  movel([0.125319, -1.305667, -2.614786, -0.791936, 1.570796, 1.696115],accel_mss,speed_ms,0,blend_radius_m)
  movel([0.123866, -1.307460, -2.613698, -0.791230, 1.570796, 1.694663],accel_mss,speed_ms,0,blend_radius_m)
  movel([0.121238, -1.311144, -2.611452, -0.789794, 1.570796, 1.692034],accel_mss,speed_ms,0,blend_radius_m)
  movel([0.120065, -1.313039, -2.610289, -0.789062, 1.570796, 1.690862],accel_mss,speed_ms,0,blend_radius_m)
  movel([0.118018, -1.316931, -2.607885, -0.787572, 1.570796, 1.688814],accel_mss,speed_ms,0,blend_radius_m)
  movel([0.117145, -1.318934, -2.606641, -0.786814, 1.570796, 1.687942],accel_mss,speed_ms,0,blend_radius_m)
  movel([0.116379, -1.320970, -2.605370, -0.786048, 1.570796, 1.687175],accel_mss,speed_ms,0,blend_radius_m)
  movel([0.115454, -1.323887, -2.603541, -0.784961, 1.570796, 1.686251],accel_mss,speed_ms,0,blend_radius_m)
  movel([0.114703, -1.326797, -2.601704, -0.783888, 1.570796, 1.685499],accel_mss,speed_ms,0,blend_radius_m)
  movel([0.114117, -1.329682, -2.599872, -0.782835, 1.570796, 1.684914],accel_mss,speed_ms,0,blend_radius_m)
  movel([0.113685, -1.332534, -2.598050, -0.781805, 1.570796, 1.684482],accel_mss,speed_ms,0,blend_radius_m)
  movel([0.113406, -1.335329, -2.596253, -0.780807, 1.570796, 1.684202],accel_mss,speed_ms,0,blend_radius_m)
  movel([0.113271, -1.338054, -2.594492, -0.779843, 1.570796, 1.684068],accel_mss,speed_ms,0,blend_radius_m)
  movel([0.113272, -1.340695, -2.592775, -0.778919, 1.570796, 1.684069],accel_mss,speed_ms,0,blend_radius_m)
  movel([0.113405, -1.343237, -2.591113, -0.778039, 1.570796, 1.684201],accel_mss,speed_ms,0,blend_radius_m)
  movel([0.114874, -1.352772, -2.584802, -0.774815, 1.570796, 1.685670],accel_mss,speed_ms,0,blend_radius_m)
  movel([0.115989, -1.360388, -2.579670, -0.772330, 1.570796, 1.686785],accel_mss,speed_ms,0,blend_radius_m)
  movel([0.116017, -1.361138, -2.579161, -0.772090, 1.570796, 1.686813],accel_mss,speed_ms,0,blend_radius_m)
  movel([0.120926, -1.357802, -2.581422, -0.773165, 1.570796, 1.691723],accel_mss,speed_ms,0,blend_radius_m)
  movel([0.125997, -1.354721, -2.583496, -0.774171, 1.570796, 1.696793],accel_mss,speed_ms,0,blend_radius_m)
  movel([0.131197, -1.351900, -2.585385, -0.775105, 1.570796, 1.701994],accel_mss,speed_ms,0,blend_radius_m)
  movel([0.136489, -1.349339, -2.587089, -0.775961, 1.570796, 1.707286],accel_mss,speed_ms,0,blend_radius_m)
  movel([0.141835, -1.347047, -2.588606, -0.776735, 1.570796, 1.712632],accel_mss,speed_ms,0,blend_radius_m)
  movel([0.147200, -1.345021, -2.589942, -0.777426, 1.570796, 1.717996],accel_mss,speed_ms,0,blend_radius_m)
  movel([0.152545, -1.343268, -2.591093, -0.778028, 1.570796, 1.723342],accel_mss,speed_ms,0,blend_radius_m)
  movel([0.157833, -1.341785, -2.592064, -0.778541, 1.570796, 1.728629],accel_mss,speed_ms,0,blend_radius_m)
  movel([0.160299, -1.341216, -2.592435, -0.778738, 1.570796, 1.731096],accel_mss,speed_ms,0,blend_radius_m)
  movel([0.162784, -1.340774, -2.592724, -0.778892, 1.570796, 1.733580],accel_mss,speed_ms,0,blend_radius_m)
  movel([0.165263, -1.340467, -2.592923, -0.778998, 1.570796, 1.736060],accel_mss,speed_ms,0,blend_radius_m)
  movel([0.167711, -1.340305, -2.593029, -0.779055, 1.570796, 1.738507],accel_mss,speed_ms,0,blend_radius_m)
  movel([0.170105, -1.340295, -2.593036, -0.779058, 1.570796, 1.740901],accel_mss,speed_ms,0,blend_radius_m)
  movel([0.172421, -1.340447, -2.592937, -0.779005, 1.570796, 1.743217],accel_mss,speed_ms,0,blend_radius_m)
  movel([0.174636, -1.340766, -2.592729, -0.778894, 1.570796, 1.745433],accel_mss,speed_ms,0,blend_radius_m)
  movel([0.176726, -1.341259, -2.592407, -0.778723, 1.570796, 1.747522],accel_mss,speed_ms,0,blend_radius_m)
  movel([0.178667, -1.341936, -2.591965, -0.778488, 1.570796, 1.749464],accel_mss,speed_ms,0,blend_radius_m)
  movel([0.180439, -1.342801, -2.591399, -0.778189, 1.570796, 1.751235],accel_mss,speed_ms,0,blend_radius_m)
  movel([0.182015, -1.343863, -2.590703, -0.777823, 1.570796, 1.752811],accel_mss,speed_ms,0,blend_radius_m)
  movel([0.183374, -1.345125, -2.589873, -0.777390, 1.570796, 1.754170],accel_mss,speed_ms,0,blend_radius_m)
  movel([0.184492, -1.346595, -2.588905, -0.776889, 1.570796, 1.755289],accel_mss,speed_ms,0,blend_radius_m)
  movel([0.185353, -1.348277, -2.587793, -0.776319, 1.570796, 1.756149],accel_mss,speed_ms,0,blend_radius_m)
  movel([0.185931, -1.350176, -2.586533, -0.775680, 1.570796, 1.756728],accel_mss,speed_ms,0,blend_radius_m)
  movel([0.186205, -1.352297, -2.585119, -0.774972, 1.570796, 1.757002],accel_mss,speed_ms,0,blend_radius_m)
  movel([0.186151, -1.355276, -2.583124, -0.773989, 1.570796, 1.756947],accel_mss,speed_ms,0,blend_radius_m)
  movel([0.185726, -1.358424, -2.581001, -0.772963, 1.570796, 1.756523],accel_mss,speed_ms,0,blend_radius_m)
  movel([0.184990, -1.361689, -2.578786, -0.771914, 1.570796, 1.755786],accel_mss,speed_ms,0,blend_radius_m)
  movel([0.184002, -1.365022, -2.576509, -0.770858, 1.570796, 1.754798],accel_mss,speed_ms,0,blend_radius_m)
  movel([0.182819, -1.368372, -2.574204, -0.769813, 1.570796, 1.753615],accel_mss,speed_ms,0,blend_radius_m)
  movel([0.181495, -1.371694, -2.571903, -0.768792, 1.570796, 1.752291],accel_mss,speed_ms,0,blend_radius_m)
  movel([0.178658, -1.378063, -2.567448, -0.766878, 1.570796, 1.749455],accel_mss,speed_ms,0,blend_radius_m)
  movel([0.176687, -1.382024, -2.564648, -0.765716, 1.570796, 1.747483],accel_mss,speed_ms,0,blend_radius_m)
  movel([0.174549, -1.385880, -2.561901, -0.764608, 1.570796, 1.745346],accel_mss,speed_ms,0,blend_radius_m)
  movel([0.172265, -1.389646, -2.559198, -0.763545, 1.570796, 1.743062],accel_mss,speed_ms,0,blend_radius_m)
  movel([0.169850, -1.393345, -2.556522, -0.762522, 1.570796, 1.740646],accel_mss,speed_ms,0,blend_radius_m)
  movel([0.167323, -1.396990, -2.553866, -0.761533, 1.570796, 1.738120],accel_mss,speed_ms,0,blend_radius_m)
  movel([0.164703, -1.400600, -2.551217, -0.760572, 1.570796, 1.735499],accel_mss,speed_ms,0,blend_radius_m)
  movel([0.159243, -1.407786, -2.545886, -0.758717, 1.570796, 1.730039],accel_mss,speed_ms,0,blend_radius_m)
  movel([0.162416, -1.409703, -2.544451, -0.758235, 1.570796, 1.733213],accel_mss,speed_ms,0,blend_radius_m)
  movel([0.164019, -1.410829, -2.543606, -0.757954, 1.570796, 1.734815],accel_mss,speed_ms,0,blend_radius_m)
  movel([0.165312, -1.412098, -2.542651, -0.757640, 1.570796, 1.736108],accel_mss,speed_ms,0,blend_radius_m)
  movel([0.165766, -1.412796, -2.542125, -0.757468, 1.570796, 1.736562],accel_mss,speed_ms,0,blend_radius_m)
  movel([0.166050, -1.413541, -2.541562, -0.757286, 1.570796, 1.736847],accel_mss,speed_ms,0,blend_radius_m)
  movel([0.166139, -1.414334, -2.540963, -0.757092, 1.570796, 1.736935],accel_mss,speed_ms,0,blend_radius_m)
  movel([0.166002, -1.415178, -2.540323, -0.756887, 1.570796, 1.736798],accel_mss,speed_ms,0,blend_radius_m)
  movel([0.165610, -1.416074, -2.539643, -0.756671, 1.570796, 1.736406],accel_mss,speed_ms,0,blend_radius_m)
  movel([0.164930, -1.417031, -2.538917, -0.756442, 1.570796, 1.735726],accel_mss,speed_ms,0,blend_radius_m)
  movel([0.163937, -1.418049, -2.538141, -0.756199, 1.570796, 1.734733],accel_mss,speed_ms,0,blend_radius_m)
  movel([0.162601, -1.419130, -2.537317, -0.755943, 1.570796, 1.733397],accel_mss,speed_ms,0,blend_radius_m)
  movel([0.161399, -1.419953, -2.536687, -0.755749, 1.570796, 1.732195],accel_mss,speed_ms,0,blend_radius_m)
  movel([0.160218, -1.420644, -2.536158, -0.755587, 1.570796, 1.731014],accel_mss,speed_ms,0,blend_radius_m)
  movel([0.159058, -1.421213, -2.535722, -0.755454, 1.570796, 1.729855],accel_mss,speed_ms,0,blend_radius_m)
  movel([0.156792, -1.422028, -2.535096, -0.755264, 1.570796, 1.727588],accel_mss,speed_ms,0,blend_radius_m)
  movel([0.155682, -1.422295, -2.534891, -0.755203, 1.570796, 1.726479],accel_mss,speed_ms,0,blend_radius_m)
  movel([0.153498, -1.422599, -2.534657, -0.755132, 1.570796, 1.724295],accel_mss,speed_ms,0,blend_radius_m)
  movel([0.151356, -1.422664, -2.534607, -0.755117, 1.570796, 1.722152],accel_mss,speed_ms,0,blend_radius_m)
  movel([0.149240, -1.422571, -2.534679, -0.755139, 1.570796, 1.720037],accel_mss,speed_ms,0,blend_radius_m)
  movel([0.145046, -1.422229, -2.534942, -0.755218, 1.570796, 1.715842],accel_mss,speed_ms,0,blend_radius_m)
  movel([0.142181, -1.424888, -2.532894, -0.754608, 1.570796, 1.712978],accel_mss,speed_ms,0,blend_radius_m)
  movel([0.140649, -1.426170, -2.531902, -0.754317, 1.570796, 1.711445],accel_mss,speed_ms,0,blend_radius_m)
  movel([0.139057, -1.427369, -2.530972, -0.754047, 1.570796, 1.709853],accel_mss,speed_ms,0,blend_radius_m)
  movel([0.137412, -1.428442, -2.530138, -0.753808, 1.570796, 1.708208],accel_mss,speed_ms,0,blend_radius_m)
  movel([0.135721, -1.429350, -2.529432, -0.753607, 1.570796, 1.706518],accel_mss,speed_ms,0,blend_radius_m)
  movel([0.133991, -1.430049, -2.528887, -0.753453, 1.570796, 1.704788],accel_mss,speed_ms,0,blend_radius_m)
  movel([0.132224, -1.430502, -2.528533, -0.753353, 1.570796, 1.703021],accel_mss,speed_ms,0,blend_radius_m)
  movel([0.131040, -1.430577, -2.528475, -0.753337, 1.570796, 1.701836],accel_mss,speed_ms,0,blend_radius_m)
  movel([0.130170, -1.430358, -2.528646, -0.753385, 1.570796, 1.700967],accel_mss,speed_ms,0,blend_radius_m)
  movel([0.129578, -1.429892, -2.529010, -0.753488, 1.570796, 1.700374],accel_mss,speed_ms,0,blend_radius_m)
  movel([0.129229, -1.429224, -2.529531, -0.753635, 1.570796, 1.700026],accel_mss,speed_ms,0,blend_radius_m)
  movel([0.129088, -1.428399, -2.530172, -0.753818, 1.570796, 1.699885],accel_mss,speed_ms,0,blend_radius_m)
  movel([0.129121, -1.427470, -2.530894, -0.754025, 1.570796, 1.699917],accel_mss,speed_ms,0,blend_radius_m)
  movel([0.129289, -1.426481, -2.531661, -0.754247, 1.570796, 1.700085],accel_mss,speed_ms,0,blend_radius_m)
  movel([0.129563, -1.425480, -2.532436, -0.754473, 1.570796, 1.700360],accel_mss,speed_ms,0,blend_radius_m)
  movel([0.130356, -1.423360, -2.534072, -0.754957, 1.570796, 1.701152],accel_mss,speed_ms,0,blend_radius_m)
  movel([0.131346, -1.421261, -2.535686, -0.755443, 1.570796, 1.702142],accel_mss,speed_ms,0,blend_radius_m)
  movel([0.133635, -1.417023, -2.538923, -0.756444, 1.570796, 1.704432],accel_mss,speed_ms,0,blend_radius_m)
  movel([0.129524, -1.413807, -2.541361, -0.757221, 1.570796, 1.700320],accel_mss,speed_ms,0,blend_radius_m)
  movel([0.125258, -1.410718, -2.543689, -0.757982, 1.570796, 1.696054],accel_mss,speed_ms,0,blend_radius_m)
  movel([0.121014, -1.407578, -2.546041, -0.758769, 1.570796, 1.691811],accel_mss,speed_ms,0,blend_radius_m)
  movel([0.118956, -1.405933, -2.547268, -0.759188, 1.570796, 1.689752],accel_mss,speed_ms,0,blend_radius_m)
  movel([0.116970, -1.404206, -2.548551, -0.759632, 1.570796, 1.687766],accel_mss,speed_ms,0,blend_radius_m)
  movel([0.115166, -1.402454, -2.549848, -0.760086, 1.570796, 1.685962],accel_mss,speed_ms,0,blend_radius_m)
  movel([0.113466, -1.400629, -2.551196, -0.760565, 1.570796, 1.684262],accel_mss,speed_ms,0,blend_radius_m)
  movel([0.110267, -1.396824, -2.553987, -0.761577, 1.570796, 1.681063],accel_mss,speed_ms,0,blend_radius_m)
  movel([0.107128, -1.392965, -2.556798, -0.762626, 1.570796, 1.677925],accel_mss,speed_ms,0,blend_radius_m)
  movel([0.103811, -1.389222, -2.559503, -0.763664, 1.570796, 1.674608],accel_mss,speed_ms,0,blend_radius_m)
  movel([0.102167, -1.391587, -2.557796, -0.763006, 1.570796, 1.672964],accel_mss,speed_ms,0,blend_radius_m)
  movel([0.100662, -1.393959, -2.556076, -0.762354, 1.570796, 1.671459],accel_mss,speed_ms,0,blend_radius_m)
  movel([0.099299, -1.396331, -2.554348, -0.761710, 1.570796, 1.670095],accel_mss,speed_ms,0,blend_radius_m)
  movel([0.098076, -1.398697, -2.552616, -0.761076, 1.570796, 1.668873],accel_mss,speed_ms,0,blend_radius_m)
  movel([0.096997, -1.401053, -2.550883, -0.760453, 1.570796, 1.667793],accel_mss,speed_ms,0,blend_radius_m)
  movel([0.096057, -1.403393, -2.549154, -0.759842, 1.570796, 1.666854],accel_mss,speed_ms,0,blend_radius_m)
  movel([0.095262, -1.405713, -2.547432, -0.759244, 1.570796, 1.666058],accel_mss,speed_ms,0,blend_radius_m)
  movel([0.094606, -1.408008, -2.545721, -0.758661, 1.570796, 1.665402],accel_mss,speed_ms,0,blend_radius_m)
  movel([0.094093, -1.410273, -2.544024, -0.758092, 1.570796, 1.664890],accel_mss,speed_ms,0,blend_radius_m)
  movel([0.093726, -1.412503, -2.542346, -0.757540, 1.570796, 1.664522],accel_mss,speed_ms,0,blend_radius_m)
  movel([0.093498, -1.414696, -2.540689, -0.757004, 1.570796, 1.664294],accel_mss,speed_ms,0,blend_radius_m)
  movel([0.093412, -1.416845, -2.539058, -0.756486, 1.570796, 1.664208],accel_mss,speed_ms,0,blend_radius_m)
  movel([0.093471, -1.418944, -2.537458, -0.755986, 1.570796, 1.664267],accel_mss,speed_ms,0,blend_radius_m)
  movel([0.093671, -1.420995, -2.535889, -0.755505, 1.570796, 1.664467],accel_mss,speed_ms,0,blend_radius_m)
  movel([0.094013, -1.422989, -2.534357, -0.755042, 1.570796, 1.664809],accel_mss,speed_ms,0,blend_radius_m)
  movel([0.094499, -1.424925, -2.532865, -0.754599, 1.570796, 1.665295],accel_mss,speed_ms,0,blend_radius_m)
  movel([0.095514, -1.427785, -2.530650, -0.753955, 1.570796, 1.666310],accel_mss,speed_ms,0,blend_radius_m)
  movel([0.096804, -1.430449, -2.528575, -0.753365, 1.570796, 1.667600],accel_mss,speed_ms,0,blend_radius_m)
  movel([0.098336, -1.432935, -2.526629, -0.752825, 1.570796, 1.669132],accel_mss,speed_ms,0,blend_radius_m)
  movel([0.100086, -1.435258, -2.524803, -0.752328, 1.570796, 1.670883],accel_mss,speed_ms,0,blend_radius_m)
  movel([0.102024, -1.437433, -2.523085, -0.751870, 1.570796, 1.672820],accel_mss,speed_ms,0,blend_radius_m)
  movel([0.104120, -1.439475, -2.521467, -0.751447, 1.570796, 1.674917],accel_mss,speed_ms,0,blend_radius_m)
  movel([0.106347, -1.441399, -2.519936, -0.751055, 1.570796, 1.677144],accel_mss,speed_ms,0,blend_radius_m)
  movel([0.108683, -1.443214, -2.518486, -0.750689, 1.570796, 1.679480],accel_mss,speed_ms,0,blend_radius_m)
  movel([0.113585, -1.446633, -2.515742, -0.750014, 1.570796, 1.684382],accel_mss,speed_ms,0,blend_radius_m)
  movel([0.118609, -1.449901, -2.513102, -0.749386, 1.570796, 1.689405],accel_mss,speed_ms,0,blend_radius_m)
  movel([0.122388, -1.452519, -2.510976, -0.748894, 1.570796, 1.693184],accel_mss,speed_ms,0,blend_radius_m)
  movel([0.123722, -1.453292, -2.510347, -0.748751, 1.570796, 1.694518],accel_mss,speed_ms,0,blend_radius_m)
  movel([0.126189, -1.454439, -2.509410, -0.748540, 1.570796, 1.696985],accel_mss,speed_ms,0,blend_radius_m)
  movel([0.126676, -1.454795, -2.509119, -0.748475, 1.570796, 1.697472],accel_mss,speed_ms,0,blend_radius_m)
  movel([0.127083, -1.455242, -2.508753, -0.748393, 1.570796, 1.697880],accel_mss,speed_ms,0,blend_radius_m)
  movel([0.127393, -1.455815, -2.508284, -0.748290, 1.570796, 1.698189],accel_mss,speed_ms,0,blend_radius_m)
  movel([0.127586, -1.456546, -2.507685, -0.748158, 1.570796, 1.698382],accel_mss,speed_ms,0,blend_radius_m)
  movel([0.127638, -1.457466, -2.506930, -0.747993, 1.570796, 1.698434],accel_mss,speed_ms,0,blend_radius_m)
  movel([0.127507, -1.458417, -2.506147, -0.747824, 1.570796, 1.698304],accel_mss,speed_ms,0,blend_radius_m)
  movel([0.127215, -1.459388, -2.505347, -0.747653, 1.570796, 1.698011],accel_mss,speed_ms,0,blend_radius_m)
  movel([0.126775, -1.460375, -2.504533, -0.747481, 1.570796, 1.697571],accel_mss,speed_ms,0,blend_radius_m)
  movel([0.126205, -1.461365, -2.503714, -0.747310, 1.570796, 1.697001],accel_mss,speed_ms,0,blend_radius_m)
  movel([0.124732, -1.463334, -2.502081, -0.746973, 1.570796, 1.695529],accel_mss,speed_ms,0,blend_radius_m)
  movel([0.123862, -1.464296, -2.501282, -0.746811, 1.570796, 1.694658],accel_mss,speed_ms,0,blend_radius_m)
  movel([0.121938, -1.466136, -2.499748, -0.746505, 1.570796, 1.692734],accel_mss,speed_ms,0,blend_radius_m)
  movel([0.119863, -1.467813, -2.498345, -0.746231, 1.570796, 1.690660],accel_mss,speed_ms,0,blend_radius_m)
  movel([0.117768, -1.469269, -2.497124, -0.745996, 1.570796, 1.688564],accel_mss,speed_ms,0,blend_radius_m)
  movel([0.115768, -1.470441, -2.496138, -0.745809, 1.570796, 1.686564],accel_mss,speed_ms,0,blend_radius_m)
  movel([0.112724, -1.471878, -2.494928, -0.745584, 1.570796, 1.683520],accel_mss,speed_ms,0,blend_radius_m)
  movel([0.111176, -1.472483, -2.494416, -0.745489, 1.570796, 1.681972],accel_mss,speed_ms,0,blend_radius_m)
  movel([0.109623, -1.473010, -2.493971, -0.745408, 1.570796, 1.680419],accel_mss,speed_ms,0,blend_radius_m)
  movel([0.106514, -1.473833, -2.493274, -0.745281, 1.570796, 1.677310],accel_mss,speed_ms,0,blend_radius_m)
  movel([0.103446, -1.474344, -2.492841, -0.745203, 1.570796, 1.674242],accel_mss,speed_ms,0,blend_radius_m)
  movel([0.100466, -1.474536, -2.492679, -0.745174, 1.570796, 1.671263],accel_mss,speed_ms,0,blend_radius_m)
  movel([0.097629, -1.474405, -2.492790, -0.745194, 1.570796, 1.668425],accel_mss,speed_ms,0,blend_radius_m)
  movel([0.096277, -1.474215, -2.492951, -0.745223, 1.570796, 1.667073],accel_mss,speed_ms,0,blend_radius_m)
  movel([0.093738, -1.473584, -2.493485, -0.745319, 1.570796, 1.664534],accel_mss,speed_ms,0,blend_radius_m)
  movel([0.092564, -1.473139, -2.493862, -0.745388, 1.570796, 1.663360],accel_mss,speed_ms,0,blend_radius_m)
  movel([0.091111, -1.472426, -2.494464, -0.745498, 1.570796, 1.661908],accel_mss,speed_ms,0,blend_radius_m)
  movel([0.089770, -1.471595, -2.495166, -0.745628, 1.570796, 1.660567],accel_mss,speed_ms,0,blend_radius_m)
  movel([0.088530, -1.470660, -2.495954, -0.745775, 1.570796, 1.659327],accel_mss,speed_ms,0,blend_radius_m)
  movel([0.087374, -1.469640, -2.496812, -0.745937, 1.570796, 1.658170],accel_mss,speed_ms,0,blend_radius_m)
  movel([0.085261, -1.467404, -2.498687, -0.746297, 1.570796, 1.656058],accel_mss,speed_ms,0,blend_radius_m)
  movel([0.083321, -1.465021, -2.500678, -0.746690, 1.570796, 1.654118],accel_mss,speed_ms,0,blend_radius_m)
  movel([0.081025, -1.461923, -2.503252, -0.747214, 1.570796, 1.651822],accel_mss,speed_ms,0,blend_radius_m)
  movel([0.078888, -1.458665, -2.505943, -0.747780, 1.570796, 1.649684],accel_mss,speed_ms,0,blend_radius_m)
  movel([0.076937, -1.455248, -2.508748, -0.748392, 1.570796, 1.647734],accel_mss,speed_ms,0,blend_radius_m)
  movel([0.075197, -1.451672, -2.511665, -0.749052, 1.570796, 1.645993],accel_mss,speed_ms,0,blend_radius_m)
  movel([0.073695, -1.447931, -2.514695, -0.749762, 1.570796, 1.644491],accel_mss,speed_ms,0,blend_radius_m)
  movel([0.072462, -1.444028, -2.517835, -0.750527, 1.570796, 1.643259],accel_mss,speed_ms,0,blend_radius_m)
  movel([0.071525, -1.439959, -2.521082, -0.751348, 1.570796, 1.642321],accel_mss,speed_ms,0,blend_radius_m)
  movel([0.070911, -1.435724, -2.524436, -0.752229, 1.570796, 1.641707],accel_mss,speed_ms,0,blend_radius_m)
  movel([0.070665, -1.432433, -2.527023, -0.752933, 1.570796, 1.641462],accel_mss,speed_ms,0,blend_radius_m)
  movel([0.070592, -1.428940, -2.529751, -0.753698, 1.570796, 1.641389],accel_mss,speed_ms,0,blend_radius_m)
  movel([0.070722, -1.425284, -2.532588, -0.754518, 1.570796, 1.641518],accel_mss,speed_ms,0,blend_radius_m)
  movel([0.071081, -1.421509, -2.535495, -0.755385, 1.570796, 1.641878],accel_mss,speed_ms,0,blend_radius_m)
  movel([0.071702, -1.417657, -2.538440, -0.756292, 1.570796, 1.642499],accel_mss,speed_ms,0,blend_radius_m)
  movel([0.072614, -1.413776, -2.541384, -0.757228, 1.570796, 1.643411],accel_mss,speed_ms,0,blend_radius_m)
  movel([0.073846, -1.409907, -2.544298, -0.758184, 1.570796, 1.644643],accel_mss,speed_ms,0,blend_radius_m)
  movel([0.074593, -1.407992, -2.545732, -0.758665, 1.570796, 1.645390],accel_mss,speed_ms,0,blend_radius_m)
  movel([0.075430, -1.406099, -2.547145, -0.759146, 1.570796, 1.646227],accel_mss,speed_ms,0,blend_radius_m)
  movel([0.077219, -1.402562, -2.549769, -0.760058, 1.570796, 1.648015],accel_mss,speed_ms,0,blend_radius_m)
  movel([0.079252, -1.399031, -2.552370, -0.760987, 1.570796, 1.650048],accel_mss,speed_ms,0,blend_radius_m)
  movel([0.081522, -1.395522, -2.554938, -0.761929, 1.570796, 1.652318],accel_mss,speed_ms,0,blend_radius_m)
  movel([0.084017, -1.392049, -2.557462, -0.762878, 1.570796, 1.654813],accel_mss,speed_ms,0,blend_radius_m)
  movel([0.086733, -1.388630, -2.559929, -0.763830, 1.570796, 1.657529],accel_mss,speed_ms,0,blend_radius_m)
  movel([0.089654, -1.385282, -2.562329, -0.764778, 1.570796, 1.660451],accel_mss,speed_ms,0,blend_radius_m)
  movel([0.092774, -1.382022, -2.564650, -0.765717, 1.570796, 1.663571],accel_mss,speed_ms,0,blend_radius_m)
  movel([0.096082, -1.378869, -2.566880, -0.766639, 1.570796, 1.666879],accel_mss,speed_ms,0,blend_radius_m)
  movel([0.093237, -1.371428, -2.572088, -0.768873, 1.570796, 1.664033],accel_mss,speed_ms,0,blend_radius_m)
  movel([0.091807, -1.367682, -2.574680, -0.770027, 1.570796, 1.662604],accel_mss,speed_ms,0,blend_radius_m)
  movel([0.090551, -1.363811, -2.577338, -0.771240, 1.570796, 1.661347],accel_mss,speed_ms,0,blend_radius_m)
  movel([0.089861, -1.360771, -2.579410, -0.772207, 1.570796, 1.660658],accel_mss,speed_ms,0,blend_radius_m)
  movel([0.089468, -1.357569, -2.581580, -0.773241, 1.570796, 1.660264],accel_mss,speed_ms,0,blend_radius_m)
  movel([0.089356, -1.354220, -2.583833, -0.774336, 1.570796, 1.660152],accel_mss,speed_ms,0,blend_radius_m)
  movel([0.089518, -1.350735, -2.586161, -0.775493, 1.570796, 1.660314],accel_mss,speed_ms,0,blend_radius_m)
  movel([0.089943, -1.347131, -2.588551, -0.776707, 1.570796, 1.660739],accel_mss,speed_ms,0,blend_radius_m)
  movel([0.090622, -1.343422, -2.590992, -0.777975, 1.570796, 1.661418],accel_mss,speed_ms,0,blend_radius_m)
  movel([0.091545, -1.339621, -2.593474, -0.779294, 1.570796, 1.662341],accel_mss,speed_ms,0,blend_radius_m)
  movel([0.092699, -1.335746, -2.595984, -0.780659, 1.570796, 1.663495],accel_mss,speed_ms,0,blend_radius_m)
  movel([0.094076, -1.331815, -2.598510, -0.782064, 1.570796, 1.664872],accel_mss,speed_ms,0,blend_radius_m)
  movel([0.095667, -1.327839, -2.601044, -0.783507, 1.570796, 1.666463],accel_mss,speed_ms,0,blend_radius_m)
  movel([0.097460, -1.323837, -2.603572, -0.784980, 1.570796, 1.668256],accel_mss,speed_ms,0,blend_radius_m)
  movel([0.099441, -1.319828, -2.606084, -0.786477, 1.570796, 1.670237],accel_mss,speed_ms,0,blend_radius_m)
  movel([0.101601, -1.315830, -2.608567, -0.787992, 1.570796, 1.672398],accel_mss,speed_ms,0,blend_radius_m)
  movel([0.103924, -1.311864, -2.611010, -0.789515, 1.570796, 1.674720],accel_mss,speed_ms,0,blend_radius_m)
  movel([0.106403, -1.307946, -2.613403, -0.791040, 1.570796, 1.677199],accel_mss,speed_ms,0,blend_radius_m)
  movel([0.109019, -1.304096, -2.615735, -0.792558, 1.570796, 1.679815],accel_mss,speed_ms,0,blend_radius_m)
  movel([0.114230, -1.296950, -2.620012, -0.795426, 1.570796, 1.685027],accel_mss,speed_ms,0,blend_radius_m)
  movel([0.117008, -1.293392, -2.622118, -0.796879, 1.570796, 1.687804],accel_mss,speed_ms,0,blend_radius_m)
  movel([0.119919, -1.289870, -2.624186, -0.798333, 1.570796, 1.690716],accel_mss,speed_ms,0,blend_radius_m)
  movel([0.122983, -1.286409, -2.626202, -0.799777, 1.570796, 1.693780],accel_mss,speed_ms,0,blend_radius_m)
  movel([0.126210, -1.283037, -2.628153, -0.801199, 1.570796, 1.697007],accel_mss,speed_ms,0,blend_radius_m)
  movel([0.129616, -1.279774, -2.630027, -0.802588, 1.570796, 1.700412],accel_mss,speed_ms,0,blend_radius_m)
  movel([0.133215, -1.276648, -2.631809, -0.803932, 1.570796, 1.704012],accel_mss,speed_ms,0,blend_radius_m)
  movel([0.137409, -1.273354, -2.633675, -0.805361, 1.570796, 1.708205],accel_mss,speed_ms,0,blend_radius_m)
  movel([0.141762, -1.270241, -2.635425, -0.806723, 1.570796, 1.712559],accel_mss,speed_ms,0,blend_radius_m)
  movel([0.146253, -1.267314, -2.637060, -0.808015, 1.570796, 1.717049],accel_mss,speed_ms,0,blend_radius_m)
  movel([0.150858, -1.264583, -2.638576, -0.809230, 1.570796, 1.721654],accel_mss,speed_ms,0,blend_radius_m)
  movel([0.155552, -1.262058, -2.639969, -0.810362, 1.570796, 1.726348],accel_mss,speed_ms,0,blend_radius_m)
  movel([0.160309, -1.259747, -2.641238, -0.811404, 1.570796, 1.731106],accel_mss,speed_ms,0,blend_radius_m)
  movel([0.165110, -1.257656, -2.642380, -0.812353, 1.570796, 1.735907],accel_mss,speed_ms,0,blend_radius_m)
  movel([0.169925, -1.255795, -2.643392, -0.813202, 1.570796, 1.740722],accel_mss,speed_ms,0,blend_radius_m)
  movel([0.174731, -1.254172, -2.644271, -0.813945, 1.570796, 1.745528],accel_mss,speed_ms,0,blend_radius_m)
  movel([0.179499, -1.252790, -2.645017, -0.814581, 1.570796, 1.750296],accel_mss,speed_ms,0,blend_radius_m)
  movel([0.184208, -1.251660, -2.645626, -0.815103, 1.570796, 1.755004],accel_mss,speed_ms,0,blend_radius_m)
  movel([0.188832, -1.250783, -2.646097, -0.815509, 1.570796, 1.759628],accel_mss,speed_ms,0,blend_radius_m)
  movel([0.193342, -1.250166, -2.646428, -0.815795, 1.570796, 1.764138],accel_mss,speed_ms,0,blend_radius_m)
  movel([0.197718, -1.249811, -2.646619, -0.815960, 1.570796, 1.768514],accel_mss,speed_ms,0,blend_radius_m)
  movel([0.201934, -1.249722, -2.646666, -0.816001, 1.570796, 1.772731],accel_mss,speed_ms,0,blend_radius_m)
  movel([0.205969, -1.249903, -2.646569, -0.815917, 1.570796, 1.776765],accel_mss,speed_ms,0,blend_radius_m)
  movel([0.210114, -1.250318, -2.646347, -0.815724, 1.570796, 1.780911],accel_mss,speed_ms,0,blend_radius_m)
  movel([0.214149, -1.250923, -2.646022, -0.815444, 1.570796, 1.784946],accel_mss,speed_ms,0,blend_radius_m)
  movel([0.218032, -1.251763, -2.645571, -0.815055, 1.570796, 1.788828],accel_mss,speed_ms,0,blend_radius_m)
  movel([0.221717, -1.252889, -2.644964, -0.814536, 1.570796, 1.792514],accel_mss,speed_ms,0,blend_radius_m)
  movel([0.225740, -1.254605, -2.644037, -0.813747, 1.570796, 1.796537],accel_mss,speed_ms,0,blend_radius_m)
  movel([0.229485, -1.256739, -2.642879, -0.812771, 1.570796, 1.800282],accel_mss,speed_ms,0,blend_radius_m)
  movel([0.232919, -1.259258, -2.641506, -0.811626, 1.570796, 1.803716],accel_mss,speed_ms,0,blend_radius_m)
  movel([0.236012, -1.262130, -2.639930, -0.810329, 1.570796, 1.806808],accel_mss,speed_ms,0,blend_radius_m)
  movel([0.238737, -1.265321, -2.638167, -0.808901, 1.570796, 1.809533],accel_mss,speed_ms,0,blend_radius_m)
  movel([0.241067, -1.268796, -2.636233, -0.807359, 1.570796, 1.811863],accel_mss,speed_ms,0,blend_radius_m)
  movel([0.242979, -1.272519, -2.634145, -0.805725, 1.570796, 1.813775],accel_mss,speed_ms,0,blend_radius_m)
  movel([0.244451, -1.276457, -2.631918, -0.804014, 1.570796, 1.815247],accel_mss,speed_ms,0,blend_radius_m)
  movel([0.246837, -1.284484, -2.627318, -0.800587, 1.570796, 1.817633],accel_mss,speed_ms,0,blend_radius_m)
  movel([0.247813, -1.288567, -2.624947, -0.798875, 1.570796, 1.818609],accel_mss,speed_ms,0,blend_radius_m)
  movel([0.248532, -1.292838, -2.622444, -0.797107, 1.570796, 1.819329],accel_mss,speed_ms,0,blend_radius_m)
  movel([0.249626, -1.300060, -2.618159, -0.794170, 1.570796, 1.820422],accel_mss,speed_ms,0,blend_radius_m)
  movel([0.250380, -1.303594, -2.616038, -0.792757, 1.570796, 1.821177],accel_mss,speed_ms,0,blend_radius_m)
  movel([0.251341, -1.306993, -2.613982, -0.791414, 1.570796, 1.822138],accel_mss,speed_ms,0,blend_radius_m)
  movel([0.252568, -1.310199, -2.612029, -0.790160, 1.570796, 1.823365],accel_mss,speed_ms,0,blend_radius_m)
  movel([0.254106, -1.313152, -2.610219, -0.789018, 1.570796, 1.824903],accel_mss,speed_ms,0,blend_radius_m)
  movel([0.256014, -1.315797, -2.608588, -0.788004, 1.570796, 1.826811],accel_mss,speed_ms,0,blend_radius_m)
  movel([0.258340, -1.318074, -2.607176, -0.787139, 1.570796, 1.829137],accel_mss,speed_ms,0,blend_radius_m)
  movel([0.259433, -1.318835, -2.606703, -0.786851, 1.570796, 1.830229],accel_mss,speed_ms,0,blend_radius_m)
  movel([0.260705, -1.319380, -2.606363, -0.786646, 1.570796, 1.831502],accel_mss,speed_ms,0,blend_radius_m)
  movel([0.261412, -1.319523, -2.606274, -0.786592, 1.570796, 1.832208],accel_mss,speed_ms,0,blend_radius_m)
  movel([0.262164, -1.319556, -2.606254, -0.786580, 1.570796, 1.832961],accel_mss,speed_ms,0,blend_radius_m)
  movel([0.262966, -1.319459, -2.606314, -0.786616, 1.570796, 1.833762],accel_mss,speed_ms,0,blend_radius_m)
  movel([0.263813, -1.319209, -2.606470, -0.786710, 1.570796, 1.834609],accel_mss,speed_ms,0,blend_radius_m)
  movel([0.264694, -1.318799, -2.606725, -0.786865, 1.570796, 1.835490],accel_mss,speed_ms,0,blend_radius_m)
  movel([0.265545, -1.318262, -2.607059, -0.787068, 1.570796, 1.836341],accel_mss,speed_ms,0,blend_radius_m)
  movel([0.267125, -1.316939, -2.607881, -0.787570, 1.570796, 1.837922],accel_mss,speed_ms,0,blend_radius_m)
  movel([0.268114, -1.315907, -2.608519, -0.787962, 1.570796, 1.838910],accel_mss,speed_ms,0,blend_radius_m)
  movel([0.268998, -1.314830, -2.609185, -0.788374, 1.570796, 1.839794],accel_mss,speed_ms,0,blend_radius_m)
  movel([0.270479, -1.312568, -2.610578, -0.789243, 1.570796, 1.841275],accel_mss,speed_ms,0,blend_radius_m)
  movel([0.271610, -1.310203, -2.612027, -0.790159, 1.570796, 1.842406],accel_mss,speed_ms,0,blend_radius_m)
  movel([0.272440, -1.307783, -2.613502, -0.791104, 1.570796, 1.843236],accel_mss,speed_ms,0,blend_radius_m)
  movel([0.273010, -1.305367, -2.614967, -0.792055, 1.570796, 1.843807],accel_mss,speed_ms,0,blend_radius_m)
  movel([0.273367, -1.303004, -2.616393, -0.792992, 1.570796, 1.844164],accel_mss,speed_ms,0,blend_radius_m)
  movel([0.273554, -1.300748, -2.617748, -0.793894, 1.570796, 1.844350],accel_mss,speed_ms,0,blend_radius_m)
  movel([0.273539, -1.296347, -2.620370, -0.795672, 1.570796, 1.844336],accel_mss,speed_ms,0,blend_radius_m)
  movel([0.273284, -1.294113, -2.621692, -0.796584, 1.570796, 1.844081],accel_mss,speed_ms,0,blend_radius_m)
  movel([0.272852, -1.291961, -2.622960, -0.797468, 1.570796, 1.843648],accel_mss,speed_ms,0,blend_radius_m)
  movel([0.272239, -1.289909, -2.624163, -0.798317, 1.570796, 1.843036],accel_mss,speed_ms,0,blend_radius_m)
  movel([0.271446, -1.287962, -2.625299, -0.799127, 1.570796, 1.842243],accel_mss,speed_ms,0,blend_radius_m)
  movel([0.270473, -1.286137, -2.626360, -0.799891, 1.570796, 1.841269],accel_mss,speed_ms,0,blend_radius_m)
  movel([0.269324, -1.284442, -2.627342, -0.800605, 1.570796, 1.840120],accel_mss,speed_ms,0,blend_radius_m)
  movel([0.267995, -1.282890, -2.628238, -0.801261, 1.570796, 1.838791],accel_mss,speed_ms,0,blend_radius_m)
  speed_ms = 0.005
  movel([0.267995, -1.273740, -2.623791, -0.814858, 1.570796, 1.838791],accel_mss,speed_ms,0,blend_radius_m)
  speed_ms = 0.040
  movel([0.263666, -1.292423, -2.612949, -0.807017, 1.570796, 1.834463],accel_mss,speed_ms,0,blend_radius_m)
  speed_ms = 0.005
  movel([0.263666, -1.301474, -2.617312, -0.793603, 1.570796, 1.834463],accel_mss,speed_ms,0,blend_radius_m)
  speed_ms = 0.025
  movel([0.261910, -1.299792, -2.618319, -0.794278, 1.570796, 1.832707],accel_mss,speed_ms,0,blend_radius_m)
  movel([0.259857, -1.298395, -2.619153, -0.794841, 1.570796, 1.830654],accel_mss,speed_ms,0,blend_radius_m)
  movel([0.258681, -1.297884, -2.619457, -0.795048, 1.570796, 1.829477],accel_mss,speed_ms,0,blend_radius_m)
  movel([0.257388, -1.297543, -2.619660, -0.795186, 1.570796, 1.828184],accel_mss,speed_ms,0,blend_radius_m)
  movel([0.255964, -1.297405, -2.619742, -0.795242, 1.570796, 1.826761],accel_mss,speed_ms,0,blend_radius_m)
  movel([0.254395, -1.297499, -2.619686, -0.795204, 1.570796, 1.825192],accel_mss,speed_ms,0,blend_radius_m)
  speed_ms = 0.005
  movel([0.254395, -1.288427, -2.615305, -0.808658, 1.570796, 1.825192],accel_mss,speed_ms,0,blend_radius_m)
  speed_ms = 0.040
  movel([0.260036, -1.283648, -2.618095, -0.810646, 1.570796, 1.830832],accel_mss,speed_ms,0,blend_radius_m)
  speed_ms = 0.005
  movel([0.260036, -1.292746, -2.622498, -0.797145, 1.570796, 1.830832],accel_mss,speed_ms,0,blend_radius_m)
  speed_ms = 0.025
  movel([0.260497, -1.290272, -2.623950, -0.798166, 1.570796, 1.831293],accel_mss,speed_ms,0,blend_radius_m)
  movel([0.260472, -1.288002, -2.625276, -0.799111, 1.570796, 1.831268],accel_mss,speed_ms,0,blend_radius_m)
  movel([0.259989, -1.285970, -2.626457, -0.799962, 1.570796, 1.830785],accel_mss,speed_ms,0,blend_radius_m)
  movel([0.259068, -1.284226, -2.627467, -0.800696, 1.570796, 1.829864],accel_mss,speed_ms,0,blend_radius_m)
  movel([0.257736, -1.282810, -2.628284, -0.801295, 1.570796, 1.828533],accel_mss,speed_ms,0,blend_radius_m)
  movel([0.256022, -1.281766, -2.628884, -0.801738, 1.570796, 1.826819],accel_mss,speed_ms,0,blend_radius_m)
  movel([0.253954, -1.281136, -2.629246, -0.802007, 1.570796, 1.824751],accel_mss,speed_ms,0,blend_radius_m)
  movel([0.252795, -1.280990, -2.629330, -0.802069, 1.570796, 1.823591],accel_mss,speed_ms,0,blend_radius_m)
  movel([0.251559, -1.280960, -2.629347, -0.802082, 1.570796, 1.822356],accel_mss,speed_ms,0,blend_radius_m)
  speed_ms = 0.005
  movel([0.251559, -1.271800, -2.624891, -0.815697, 1.570796, 1.822356],accel_mss,speed_ms,0,blend_radius_m)
  speed_ms = 0.040
  movel([0.258347, -1.267761, -2.627169, -0.817459, 1.570796, 1.829143],accel_mss,speed_ms,0,blend_radius_m)
  speed_ms = 0.005
  movel([0.258347, -1.276941, -2.631643, -0.803805, 1.570796, 1.829143],accel_mss,speed_ms,0,blend_radius_m)
  speed_ms = 0.025
  movel([0.258384, -1.275747, -2.632321, -0.804321, 1.570796, 1.829181],accel_mss,speed_ms,0,blend_radius_m)
  movel([0.258271, -1.274594, -2.632974, -0.804821, 1.570796, 1.829067],accel_mss,speed_ms,0,blend_radius_m)
  movel([0.257621, -1.272434, -2.634193, -0.805762, 1.570796, 1.828417],accel_mss,speed_ms,0,blend_radius_m)
  movel([0.256463, -1.270524, -2.635267, -0.806599, 1.570796, 1.827259],accel_mss,speed_ms,0,blend_radius_m)
  movel([0.254866, -1.268928, -2.636160, -0.807301, 1.570796, 1.825663],accel_mss,speed_ms,0,blend_radius_m)
  movel([0.252900, -1.267700, -2.636845, -0.807844, 1.570796, 1.823697],accel_mss,speed_ms,0,blend_radius_m)
  movel([0.250644, -1.266901, -2.637290, -0.808198, 1.570796, 1.821440],accel_mss,speed_ms,0,blend_radius_m)
  movel([0.249426, -1.266682, -2.637412, -0.808296, 1.570796, 1.820222],accel_mss,speed_ms,0,blend_radius_m)
  movel([0.246869, -1.266632, -2.637439, -0.808318, 1.570796, 1.817665],accel_mss,speed_ms,0,blend_radius_m)
  movel([0.245547, -1.266815, -2.637338, -0.808237, 1.570796, 1.816343],accel_mss,speed_ms,0,blend_radius_m)
  speed_ms = 0.005
  movel([0.245547, -1.257584, -2.632818, -0.821986, 1.570796, 1.816343],accel_mss,speed_ms,0,blend_radius_m)
  speed_ms = 0.040
  movel([0.254982, -1.253067, -2.635286, -0.824036, 1.570796, 1.825778],accel_mss,speed_ms,0,blend_radius_m)
  speed_ms = 0.005
  movel([0.254982, -1.262319, -2.639825, -0.810244, 1.570796, 1.825778],accel_mss,speed_ms,0,blend_radius_m)
  speed_ms = 0.025
  movel([0.253875, -1.260016, -2.641091, -0.811283, 1.570796, 1.824671],accel_mss,speed_ms,0,blend_radius_m)
  movel([0.252359, -1.258018, -2.642183, -0.812188, 1.570796, 1.823155],accel_mss,speed_ms,0,blend_radius_m)
  movel([0.250459, -1.256389, -2.643069, -0.812930, 1.570796, 1.821255],accel_mss,speed_ms,0,blend_radius_m)
  movel([0.248193, -1.255176, -2.643728, -0.813485, 1.570796, 1.818989],accel_mss,speed_ms,0,blend_radius_m)
  movel([0.245585, -1.254440, -2.644126, -0.813823, 1.570796, 1.816382],accel_mss,speed_ms,0,blend_radius_m)
  movel([0.244162, -1.254265, -2.644221, -0.813903, 1.570796, 1.814958],accel_mss,speed_ms,0,blend_radius_m)
  movel([0.242664, -1.254228, -2.644241, -0.813920, 1.570796, 1.813461],accel_mss,speed_ms,0,blend_radius_m)
  movel([0.241092, -1.254336, -2.644183, -0.813870, 1.570796, 1.811889],accel_mss,speed_ms,0,blend_radius_m)
  movel([0.239450, -1.254595, -2.644043, -0.813752, 1.570796, 1.810246],accel_mss,speed_ms,0,blend_radius_m)
  movel([0.237745, -1.255008, -2.643819, -0.813562, 1.570796, 1.808541],accel_mss,speed_ms,0,blend_radius_m)
  movel([0.235979, -1.255583, -2.643507, -0.813299, 1.570796, 1.806775],accel_mss,speed_ms,0,blend_radius_m)
  speed_ms = 0.005
  movel([0.235979, -1.246300, -2.638937, -0.827152, 1.570796, 1.806775],accel_mss,speed_ms,0,blend_radius_m)
  speed_ms = 0.040
  movel([0.246368, -1.239972, -2.642302, -0.830115, 1.570796, 1.817164],accel_mss,speed_ms,0,blend_radius_m)
  speed_ms = 0.005
  movel([0.246368, -1.249284, -2.646901, -0.816205, 1.570796, 1.817164],accel_mss,speed_ms,0,blend_radius_m)
  speed_ms = 0.025
  movel([0.246209, -1.247542, -2.647830, -0.817016, 1.570796, 1.817005],accel_mss,speed_ms,0,blend_radius_m)
  movel([0.245760, -1.245957, -2.648673, -0.817758, 1.570796, 1.816557],accel_mss,speed_ms,0,blend_radius_m)
  movel([0.245031, -1.244559, -2.649414, -0.818415, 1.570796, 1.815827],accel_mss,speed_ms,0,blend_radius_m)
  movel([0.244031, -1.243382, -2.650037, -0.818970, 1.570796, 1.814828],accel_mss,speed_ms,0,blend_radius_m)
  movel([0.242506, -1.242272, -2.650622, -0.819495, 1.570796, 1.813302],accel_mss,speed_ms,0,blend_radius_m)
  movel([0.240726, -1.241447, -2.651056, -0.819886, 1.570796, 1.811523],accel_mss,speed_ms,0,blend_radius_m)
  movel([0.238414, -1.240758, -2.651418, -0.820213, 1.570796, 1.809211],accel_mss,speed_ms,0,blend_radius_m)
  movel([0.235892, -1.240398, -2.651607, -0.820384, 1.570796, 1.806688],accel_mss,speed_ms,0,blend_radius_m)
  movel([0.233181, -1.240413, -2.651599, -0.820377, 1.570796, 1.803977],accel_mss,speed_ms,0,blend_radius_m)
  movel([0.230303, -1.240852, -2.651369, -0.820168, 1.570796, 1.801100],accel_mss,speed_ms,0,blend_radius_m)
  movel([0.227293, -1.241765, -2.650889, -0.819735, 1.570796, 1.798090],accel_mss,speed_ms,0,blend_radius_m)
  movel([0.225769, -1.242400, -2.650555, -0.819434, 1.570796, 1.796565],accel_mss,speed_ms,0,blend_radius_m)
  movel([0.222755, -1.244014, -2.649703, -0.818672, 1.570796, 1.793551],accel_mss,speed_ms,0,blend_radius_m)
  movel([0.221293, -1.244982, -2.649191, -0.818216, 1.570796, 1.792090],accel_mss,speed_ms,0,blend_radius_m)
  movel([0.219885, -1.246057, -2.648621, -0.817712, 1.570796, 1.790681],accel_mss,speed_ms,0,blend_radius_m)
  movel([0.218541, -1.247233, -2.647995, -0.817161, 1.570796, 1.789338],accel_mss,speed_ms,0,blend_radius_m)
  speed_ms = 0.005
  movel([0.218541, -1.237913, -2.643387, -0.831089, 1.570796, 1.789338],accel_mss,speed_ms,0,blend_radius_m)
  speed_ms = 0.040
  movel([0.230645, -1.226985, -2.649062, -0.836342, 1.570796, 1.801442],accel_mss,speed_ms,0,blend_radius_m)
  speed_ms = 0.005
  movel([0.230645, -1.236352, -2.653719, -0.822318, 1.570796, 1.801442],accel_mss,speed_ms,0,blend_radius_m)
  speed_ms = 0.025
  movel([0.227546, -1.235639, -2.654089, -0.822660, 1.570796, 1.798342],accel_mss,speed_ms,0,blend_radius_m)
  movel([0.224143, -1.235327, -2.654251, -0.822811, 1.570796, 1.794939],accel_mss,speed_ms,0,blend_radius_m)
  movel([0.220507, -1.235475, -2.654175, -0.822740, 1.570796, 1.791303],accel_mss,speed_ms,0,blend_radius_m)
  movel([0.218626, -1.235735, -2.654039, -0.822614, 1.570796, 1.789422],accel_mss,speed_ms,0,blend_radius_m)
  movel([0.216714, -1.236132, -2.653833, -0.822423, 1.570796, 1.787510],accel_mss,speed_ms,0,blend_radius_m)
  movel([0.214784, -1.236670, -2.653554, -0.822165, 1.570796, 1.785580],accel_mss,speed_ms,0,blend_radius_m)
  movel([0.212846, -1.237354, -2.653198, -0.821837, 1.570796, 1.783643],accel_mss,speed_ms,0,blend_radius_m)
  movel([0.210909, -1.238190, -2.652762, -0.821437, 1.570796, 1.781705],accel_mss,speed_ms,0,blend_radius_m)
  movel([0.208981, -1.239187, -2.652241, -0.820961, 1.570796, 1.779778],accel_mss,speed_ms,0,blend_radius_m)
  movel([0.207073, -1.240346, -2.651634, -0.820409, 1.570796, 1.777869],accel_mss,speed_ms,0,blend_radius_m)
  movel([0.205198, -1.241676, -2.650936, -0.819777, 1.570796, 1.775994],accel_mss,speed_ms,0,blend_radius_m)
  movel([0.203363, -1.243178, -2.650145, -0.819066, 1.570796, 1.774159],accel_mss,speed_ms,0,blend_radius_m)
  movel([0.201579, -1.244861, -2.649255, -0.818273, 1.570796, 1.772376],accel_mss,speed_ms,0,blend_radius_m)
  speed_ms = 0.005
  movel([0.201579, -1.235530, -2.644636, -0.832223, 1.570796, 1.772376],accel_mss,speed_ms,0,blend_radius_m)
  speed_ms = 0.040
  movel([0.211540, -1.222257, -2.651475, -0.838657, 1.570796, 1.782336],accel_mss,speed_ms,0,blend_radius_m)
  speed_ms = 0.005
  movel([0.211540, -1.231642, -2.656154, -0.824593, 1.570796, 1.782336],accel_mss,speed_ms,0,blend_radius_m)
  speed_ms = 0.025
  movel([0.209893, -1.231427, -2.656265, -0.824698, 1.570796, 1.780689],accel_mss,speed_ms,0,blend_radius_m)
  movel([0.208146, -1.231395, -2.656281, -0.824713, 1.570796, 1.778942],accel_mss,speed_ms,0,blend_radius_m)
  movel([0.206318, -1.231551, -2.656201, -0.824637, 1.570796, 1.777114],accel_mss,speed_ms,0,blend_radius_m)
  movel([0.204427, -1.231884, -2.656029, -0.824476, 1.570796, 1.775223],accel_mss,speed_ms,0,blend_radius_m)
  movel([0.202487, -1.232393, -2.655767, -0.824228, 1.570796, 1.773284],accel_mss,speed_ms,0,blend_radius_m)
  movel([0.200520, -1.233075, -2.655416, -0.823898, 1.570796, 1.771316],accel_mss,speed_ms,0,blend_radius_m)
  movel([0.198544, -1.233921, -2.654979, -0.823489, 1.570796, 1.769341],accel_mss,speed_ms,0,blend_radius_m)
  movel([0.196572, -1.234929, -2.654457, -0.823003, 1.570796, 1.767369],accel_mss,speed_ms,0,blend_radius_m)
  movel([0.194628, -1.236092, -2.653854, -0.822443, 1.570796, 1.765425],accel_mss,speed_ms,0,blend_radius_m)
  movel([0.192731, -1.237395, -2.653177, -0.821818, 1.570796, 1.763527],accel_mss,speed_ms,0,blend_radius_m)
  movel([0.190896, -1.238819, -2.652434, -0.821136, 1.570796, 1.761693],accel_mss,speed_ms,0,blend_radius_m)
  movel([0.189139, -1.240353, -2.651631, -0.820405, 1.570796, 1.759936],accel_mss,speed_ms,0,blend_radius_m)
  movel([0.187475, -1.241978, -2.650777, -0.819634, 1.570796, 1.758271],accel_mss,speed_ms,0,blend_radius_m)
  movel([0.185915, -1.243685, -2.649877, -0.818827, 1.570796, 1.756712],accel_mss,speed_ms,0,blend_radius_m)
  movel([0.184484, -1.245454, -2.648941, -0.817995, 1.570796, 1.755280],accel_mss,speed_ms,0,blend_radius_m)
  movel([0.183189, -1.247270, -2.647975, -0.817143, 1.570796, 1.753985],accel_mss,speed_ms,0,blend_radius_m)
  speed_ms = 0.005
  movel([0.183189, -1.237950, -2.643367, -0.831071, 1.570796, 1.753985],accel_mss,speed_ms,0,blend_radius_m)
  speed_ms = 0.040
  movel([0.190188, -1.224714, -2.650225, -0.837451, 1.570796, 1.760985],accel_mss,speed_ms,0,blend_radius_m)
  speed_ms = 0.005
  movel([0.190188, -1.234090, -2.654892, -0.823408, 1.570796, 1.760985],accel_mss,speed_ms,0,blend_radius_m)
  speed_ms = 0.025
  movel([0.188519, -1.234013, -2.654931, -0.823444, 1.570796, 1.759315],accel_mss,speed_ms,0,blend_radius_m)
  movel([0.186727, -1.234256, -2.654806, -0.823327, 1.570796, 1.757523],accel_mss,speed_ms,0,blend_radius_m)
  movel([0.184851, -1.234786, -2.654532, -0.823072, 1.570796, 1.755647],accel_mss,speed_ms,0,blend_radius_m)
  movel([0.182918, -1.235562, -2.654129, -0.822697, 1.570796, 1.753715],accel_mss,speed_ms,0,blend_radius_m)
  movel([0.180963, -1.236553, -2.653615, -0.822221, 1.570796, 1.751760],accel_mss,speed_ms,0,blend_radius_m)
  movel([0.179021, -1.237720, -2.653007, -0.821662, 1.570796, 1.749817],accel_mss,speed_ms,0,blend_radius_m)
  movel([0.177119, -1.239023, -2.652327, -0.821039, 1.570796, 1.747915],accel_mss,speed_ms,0,blend_radius_m)
  movel([0.175294, -1.240430, -2.651590, -0.820369, 1.570796, 1.746091],accel_mss,speed_ms,0,blend_radius_m)
  movel([0.173490, -1.241972, -2.650780, -0.819637, 1.570796, 1.744286],accel_mss,speed_ms,0,blend_radius_m)
  movel([0.171762, -1.243610, -2.649916, -0.818862, 1.570796, 1.742558],accel_mss,speed_ms,0,blend_radius_m)
  movel([0.170136, -1.245330, -2.649006, -0.818053, 1.570796, 1.740932],accel_mss,speed_ms,0,blend_radius_m)
  movel([0.168650, -1.247113, -2.648059, -0.817217, 1.570796, 1.739446],accel_mss,speed_ms,0,blend_radius_m)
  movel([0.167332, -1.248938, -2.647086, -0.816366, 1.570796, 1.738129],accel_mss,speed_ms,0,blend_radius_m)
  movel([0.166213, -1.250787, -2.646095, -0.815507, 1.570796, 1.737009],accel_mss,speed_ms,0,blend_radius_m)
  movel([0.165329, -1.252644, -2.645096, -0.814649, 1.570796, 1.736126],accel_mss,speed_ms,0,blend_radius_m)
  movel([0.164705, -1.254489, -2.644100, -0.813800, 1.570796, 1.735502],accel_mss,speed_ms,0,blend_radius_m)
  speed_ms = 0.005
  movel([0.164705, -1.245201, -2.639525, -0.827663, 1.570796, 1.735502],accel_mss,speed_ms,0,blend_radius_m)
  speed_ms = 0.040
  movel([0.166778, -1.233885, -2.645495, -0.833009, 1.570796, 1.737575],accel_mss,speed_ms,0,blend_radius_m)
  speed_ms = 0.005
  movel([0.166778, -1.243223, -2.650121, -0.819045, 1.570796, 1.737575],accel_mss,speed_ms,0,blend_radius_m)
  speed_ms = 0.025
  movel([0.164066, -1.244515, -2.649438, -0.818436, 1.570796, 1.734863],accel_mss,speed_ms,0,blend_radius_m)
  movel([0.161231, -1.246176, -2.648557, -0.817656, 1.570796, 1.732028],accel_mss,speed_ms,0,blend_radius_m)
  movel([0.158422, -1.248144, -2.647509, -0.816735, 1.570796, 1.729218],accel_mss,speed_ms,0,blend_radius_m)
  movel([0.155787, -1.250356, -2.646326, -0.815707, 1.570796, 1.726583],accel_mss,speed_ms,0,blend_radius_m)
  movel([0.153469, -1.252750, -2.645039, -0.814600, 1.570796, 1.724265],accel_mss,speed_ms,0,blend_radius_m)
  movel([0.152472, -1.253998, -2.644366, -0.814026, 1.570796, 1.723269],accel_mss,speed_ms,0,blend_radius_m)
  movel([0.151611, -1.255266, -2.643679, -0.813444, 1.570796, 1.722407],accel_mss,speed_ms,0,blend_radius_m)
  movel([0.150897, -1.256553, -2.642980, -0.812856, 1.570796, 1.721694],accel_mss,speed_ms,0,blend_radius_m)
  movel([0.150350, -1.257848, -2.642275, -0.812266, 1.570796, 1.721146],accel_mss,speed_ms,0,blend_radius_m)
  movel([0.149991, -1.259141, -2.641569, -0.811679, 1.570796, 1.720787],accel_mss,speed_ms,0,blend_radius_m)
  movel([0.149830, -1.260432, -2.640862, -0.811094, 1.570796, 1.720627],accel_mss,speed_ms,0,blend_radius_m)
  speed_ms = 0.005
  movel([0.149830, -1.251172, -2.636314, -0.824903, 1.570796, 1.720627],accel_mss,speed_ms,0,blend_radius_m)
  speed_ms = 0.040
  movel([0.146520, -1.247161, -2.638475, -0.826753, 1.570796, 1.717316],accel_mss,speed_ms,0,blend_radius_m)
  speed_ms = 0.005
  movel([0.146520, -1.256440, -2.643042, -0.812907, 1.570796, 1.717316],accel_mss,speed_ms,0,blend_radius_m)
  speed_ms = 0.025
  movel([0.142921, -1.259714, -2.641256, -0.811419, 1.570796, 1.713717],accel_mss,speed_ms,0,blend_radius_m)
  movel([0.141219, -1.261464, -2.640296, -0.810629, 1.570796, 1.712016],accel_mss,speed_ms,0,blend_radius_m)
  movel([0.139650, -1.263269, -2.639302, -0.809818, 1.570796, 1.710446],accel_mss,speed_ms,0,blend_radius_m)
  movel([0.138258, -1.265126, -2.638275, -0.808988, 1.570796, 1.709055],accel_mss,speed_ms,0,blend_radius_m)
  movel([0.137089, -1.267024, -2.637221, -0.808144, 1.570796, 1.707885],accel_mss,speed_ms,0,blend_radius_m)
  movel([0.136194, -1.268951, -2.636147, -0.807291, 1.570796, 1.706990],accel_mss,speed_ms,0,blend_radius_m)
  movel([0.135613, -1.270901, -2.635055, -0.806433, 1.570796, 1.706409],accel_mss,speed_ms,0,blend_radius_m)
  speed_ms = 0.005
  # Splitting Linear movement in 2 (instruction 3386: MoveL 3110)
  movel([0.135613, -1.248262, -2.623696, -0.840431, 1.570796, 1.706409],accel_mss,speed_ms,0,blend_radius_m)
  movel([0.135613, -1.226892, -2.611993, -0.873504, 1.570796, 1.706409],accel_mss,speed_ms,0,blend_radius_m)
  speed_ms = 1.000
  movel([0.135613, -1.226892, -2.611993, -0.873504, 1.570796, 1.706409],accel_mss,speed_ms,0,blend_radius_m)
  # Splitting Linear movement in 6 (instruction 3389: MoveL 3112)
  movel([0.135613, -1.193983, -2.591775, -0.926631, 1.570796, 1.706409],accel_mss,speed_ms,0,blend_radius_m)
  movel([0.135613, -1.164289, -2.570732, -0.977368, 1.570796, 1.706409],accel_mss,speed_ms,0,blend_radius_m)
  movel([0.135613, -1.137604, -2.548935, -1.025850, 1.570796, 1.706409],accel_mss,speed_ms,0,blend_radius_m)
  movel([0.135613, -1.113724, -2.526446, -1.072219, 1.570796, 1.706409],accel_mss,speed_ms,0,blend_radius_m)
  movel([0.135613, -1.092452, -2.503317, -1.116620, 1.570796, 1.706409],accel_mss,speed_ms,0,blend_radius_m)
  movel([0.135613, -1.073596, -2.479596, -1.159197, 1.570796, 1.706409],accel_mss,speed_ms,0,blend_radius_m)
  # End of main program
end

Machining2()
